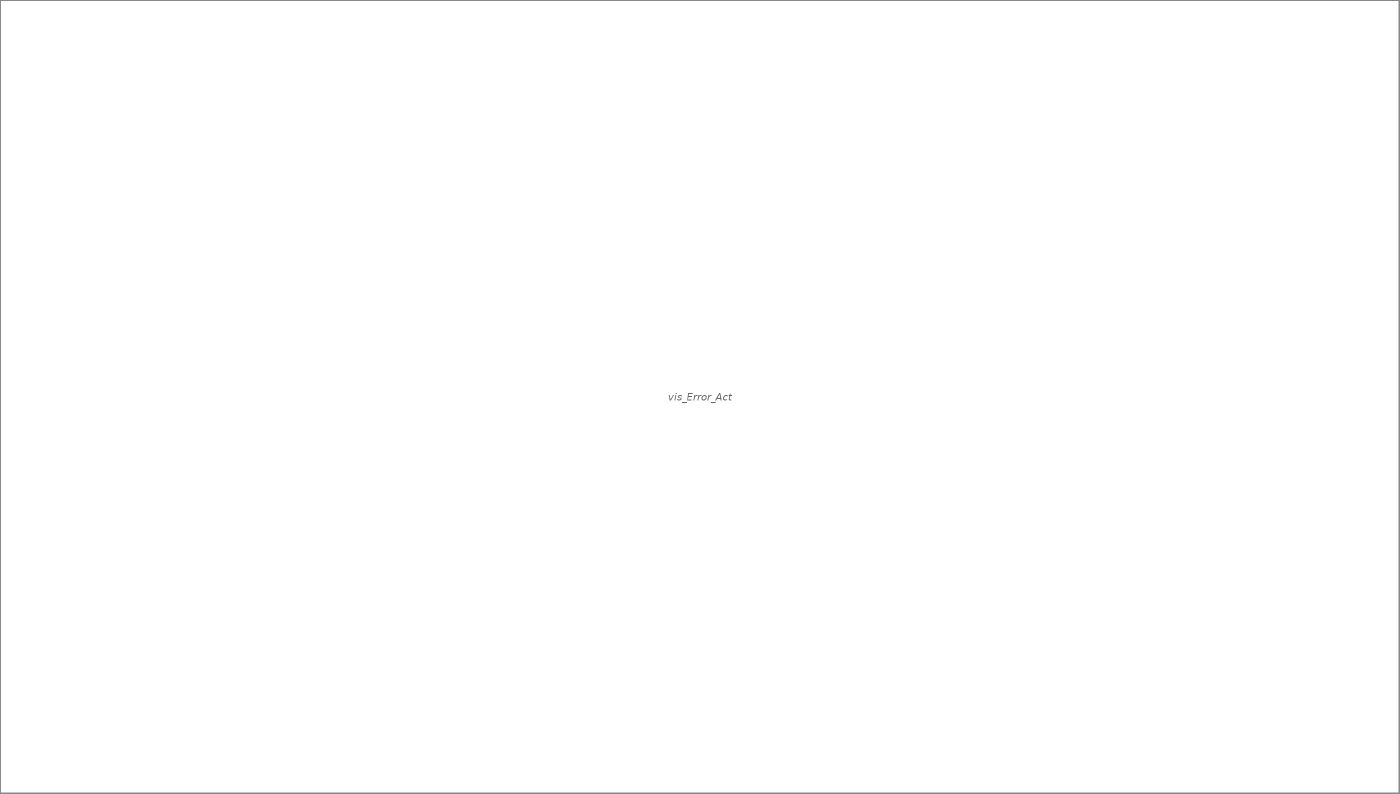
VISUALIZATION ERROR_Tab_1  // 1428x810
    TabControl (0,0 1428x810)
        shows vis_Error_Act()
        shows vis_Error_History()
        shows vis_Error_Search()
        [0]: TabTitle=Actual
        [1]: TabTitle=History
        [2]: TabTitle=Search
END_VISUALIZATION

(* stored: Version 1.1.0.1, ProductVersion 3.1.4024.13
   Visu ERROR_Tab_1: Id {d218411c-9714-4c26-ab80-d101521a00e9} *)
